Fanuc KAREL source: kd00057.KL

-- PROVISIONAL review KL for V1013-1; original PC SHA256 a089822aeba1585a45aa053b6cc0e1af705a7e464f7f30ea62bad0d778fc0552
-- Incomplete behavior may be omitted. Consult companion uncertainty JSON. Do not deploy.
PROGRAM KD00057
%NOLOCKGROUP
VAR
  I : INTEGER
  J : INTEGER
  B : BOOLEAN
  R : REAL
  S : STRING[80]
-- UNRESOLVED_DECL P type=000101
-- UNRESOLVED_DECL Q type=000101
BEGIN
  -- UNRESOLVED_PC offsets 5-37; opcodes 01,22,1C,06,22,1C,07,82,0B
  -- UNRESOLVED_PC offsets 42-46; opcodes 7F
END KD00057
